Fanuc KAREL source: KT00609.KL

PROGRAM KT00609
%NOLOCKGROUP
VAR
  R1: REAL
  R2: REAL
  OUT: BOOLEAN
BEGIN
  R1 = 2.0
  R2 = 3.0
  R1 = 2.0
  R2 = 3.0
  OUT = NOT R1
END KT00609
